TYPE ST_PLCTOROBOT :
STRUCT
	arbyOutput				:ARRAY[0..63] OF BYTE;
END_STRUCT
END_TYPE

(* stored: Version 1.1.0.1, ProductVersion 3.1.4024.15
   DUT ST_PLCTOROBOT: Id {c4501eb6-c38f-488a-abc9-497fbeac1ff3} *)
